(*
SPDX-FileCopyrightText: © 2026 Oleksandr Tiutyk <trofimich@gmail.com>
SPDX-License-Identifier: MIT
License: https://opensource.org/license/mit
*)

(*!
<summary>Enumerates a borrowed stack using an independent cursor.</summary>
<description>
The source must be non-null, outlive the cursor and remain structurally unchanged during traversal. The caller
explicitly releases a dynamically created cursor. Current is borrowed read-only data, never an ownership
transfer. Traverses from top to bottom. Supports both fixed-capacity and dynamic stacks. MoveNext stops
advancing at the end position of an unchanged source; repeated exhausted calls return FALSE until Reset.
A null constructor source is diagnosed by traversal/current access, never by FB_init.
</description>
*)

{attribute 'no_explicit_call' := 'do not call this function block directly'}
{attribute 'enable_dynamic_creation'}
FUNCTION_BLOCK StackEnumerator EXTENDS TOF_Core.Object IMPLEMENTS TOF_Core.IEnumerator
VAR_STAT
	//! <summary>Class name shared by all instances of this function block.</summary>
	{attribute 'hide'} 
	_ClassName : STRING := __POUNAME();
END_VAR
VAR
	{attribute 'hide'} 
	_Stack : IReadOnlyStack;
	{attribute 'hide'} 
	//!<summary>Top-relative position; minus one represents the cursor before the first entry.</summary>
	_CurrentIndex : DINT := -1;
	
	{attribute 'hide'} 
	_GenericValue : TOF_Core.GENERIC_VALUE;
END_VAR

(*!
<summary>Borrows the concrete cursor class name without transferring storage ownership.</summary>
*)
{attribute 'monitoring' := 'call'}
PROPERTY ClassName : REFERENCE TO STRING
GET
ClassName REF= _ClassName;
END_GET
END_PROPERTY

(*!
<summary>Exposes a read-only borrowed view of the current entry.</summary>
<description>
Reading Current before the first successful MoveNext, after Reset or after exhaustion yields an empty
descriptor. Otherwise payload is borrowed, with no disposal rights. Do not modify or release the descriptor.
The view may change on subsequent property access, cursor movement or source mutation.
Missing source raises DataMemberNotSpecifiedException before source access or cursor advancement.
</description>
*)
{attribute 'monitoring' := 'call'}
PROPERTY FINAL Current : REFERENCE TO TOF_Core.GENERIC_VALUE
GET
requireSource();

IF _CurrentIndex >= TOF_Core.SignedInt32.ZERO AND_THEN _CurrentIndex < _Stack.Length THEN
	_GenericValue := _Stack.GetByIndex(index := _CurrentIndex); 
ELSE
	_GenericValue.Reset();	
END_IF 

Current REF= _GenericValue;
END_GET
END_PROPERTY

(*!
<summary>Binds the borrowed source for enumeration.</summary>
<description>
The source must be non-null and outlive the cursor. Only the reference is assigned; no allocation, callbacks
or throwing validation are performed. A null source remains invalid configuration and is reported by
MoveNext or current-value access without throwing from initialization.
</description>
*)
METHOD FB_init : BOOL
VAR_INPUT
	bInitRetains : BOOL; // TRUE: the retain variables are initialized (reset warm / reset cold)
	bInCopyCode : BOOL;  // TRUE: the instance will be copied to the copy code afterward (online change)
	stack : IReadOnlyStack;
END_VAR
_Stack := stack;
END_METHOD

(*!
<summary>Advances the cursor to the next source position.</summary>
<description>
The source must be live, non-null and structurally unchanged during traversal. TRUE identifies a current
entry. The index advances only while below source Length and stops at the end position. Repeated exhausted
calls return FALSE without incrementing the index; reading Current yields an empty descriptor. Reset allows
traversal from the beginning again. No snapshot or mutation detection is provided. Descendants cannot override
this cursor operation; advancement, reset and borrowed current views use the same cursor state.
Missing source raises DataMemberNotSpecifiedException before source access or cursor advancement.
</description>
*)
{attribute "object_name" := "MoveNext"}
METHOD FINAL MoveNext : BOOL
requireSource();

IF _CurrentIndex < _Stack.Length THEN
	_CurrentIndex := _CurrentIndex + 1;
END_IF

MoveNext := _CurrentIndex < _Stack.Length;
END_METHOD

(*!
<summary>Provides the library namespace for diagnostics.</summary>
<description>
Borrowed read-only reference to compiler-initialized metadata; no ownership transfer.
</description>
*)
{attribute 'monitoring' := 'call'}
PROPERTY NamespaceName : REFERENCE TO STRING
GET
NamespaceName REF= CurrentNamespace.Name;
END_GET
END_PROPERTY

(*!
<summary>Places the cursor before the first source entry.</summary>
<description>
The next MoveNext starts at zero. Does not modify the source or release payload; reading Current now yields an
empty descriptor. Descendants cannot override this cursor operation; advancement, reset and borrowed current
views use the same cursor state.
</description>
*)
{attribute "object_name" := "Reset"}
METHOD FINAL Reset
_CurrentIndex := -1;
END_METHOD

(*!
<summary>Reports the size of this function-block instance.</summary>
<description>
Measured in bytes; includes inline storage but excludes separately allocated buffers, payload and enumerators.
</description>
*)
{attribute 'monitoring' := 'call'}
PROPERTY SelfSize : ULINT
GET
SelfSize := XSIZEOF(THIS^);
END_GET
END_PROPERTY

(*!
<summary>Requires the configured source before traversal or current-value access.</summary>
<description>
A missing mandatory source is configuration failure, not an empty collection. Raises a framework diagnostic
outside lifecycle methods and before mutation; it does not validate arbitrary pointer lifetime.
</description>
*)
METHOD PRIVATE requireSource
IF _Stack = 0 THEN
	TOF_Core.Exceptions.ThrowDataMemberNotSpecified(
		sourceNamespaceName := NamespaceName,
		sourceClassName := ClassName,
		sourcePOUName := __POUNAME(),
		sourcePosition := __POSITION(),
		dataMemberName := 'stack'
	);
END_IF
END_METHOD

END_FUNCTION_BLOCK

(* stored: Version 1.1.0.1
   POU StackEnumerator: Id {e416d399-9dd5-4cb2-b9ab-6df401117b4b}, SpecialFunc None
   Property ClassName: Id {26c6f006-587c-4952-acea-42d8f9ee18b5}
   Get Get: Id {625934d1-371a-449b-80c4-6fdb2abaadd7}
   Property Current: Id {7b130588-92b9-47cf-9ece-7bab9548bbf7}
   Get Get: Id {2a2cfc97-9e56-485a-990c-1429fa351b49}
   Method FB_init: Id {058de72d-67eb-4fa1-bd5e-1ce98906e144}
   Method MoveNext: Id {60bdc8b6-a79f-413f-a052-685c1b66ff7c}
   Property NamespaceName: Id {41db8516-569e-46a2-b3c2-7e7b20f0c340}
   Get Get: Id {7c548c9d-cc27-4886-9a7d-beb0d647cfc5}
   Method Reset: Id {bbc5a77c-4535-4950-b859-06b46db423a4}
   Property SelfSize: Id {c679d536-5abc-4b01-9533-75c921118918}
   Get Get: Id {e4c32193-d837-407c-aab4-c3a364acec64}
   Method requireSource: Id {95319154-56fd-4a64-b013-7fd3a687aa75} *)
